TYPE ST_PLC_To_VisuPLC :
STRUCT
	lifeBit: BOOL;
	
// General
	Description				: STRING(30);
	prodType				: E_Prod_Type;	
	RPM_FeedBack			: REAL;
	Flow_FeedBack			: REAL;
	fBlendingPercenatge		: DINT;
	
// Component
	arr_Component			: ARRAY [1..10] OF ST_Prod_Ingredient;

	iActual_Component		: INT;
	bDissolving_Active		: BOOL;
	bBlending_Active		: BOOL;
	bMainPause_Active		: BOOL;

END_STRUCT
END_TYPE

(* stored: Version 1.1.0.1, ProductVersion 3.1.4024.15
   DUT ST_PLC_To_VisuPLC: Id {4ca841ff-0e69-41d3-8667-041439910d64} *)
